Fanuc KAREL source: kb00111.KL

-- PROVISIONAL review KL for V1013-1; original PC SHA256 eba65beb3902ab2f39382df96c91639f241133c323665944e3cb6c7573fb4e1d
-- Incomplete behavior may be omitted. Consult companion uncertainty JSON. Do not deploy.
PROGRAM KB00111
%NOLOCKGROUP
BEGIN
  -- UNRESOLVED_PC offsets 5-21; opcodes 27,22,31,23
  -- UNRESOLVED_PC offsets 26-30; opcodes 7F
END KB00111
